(* IEC 61131-3 sources: nautilus/website/lessons/b4-counter/variants/bad-count-per-scan, 1 file *)

(* ---- program.st ---- *)
PROGRAM Counter
VAR n : INT; END_VAR
IF Reset THEN n := 0; ELSIF Eye THEN n := n + 1; END_IF;
Count := n;
Full := n >= 5;
END_PROGRAM
